(* IEC 61131-3 sources: model-first-plc-agent-ai/results/T3-B-12, 1 file *)

(* ---- b_code.st ---- *)
FUNCTION_BLOCK FillingTankControl
VAR_INPUT
    start : BOOL;
    stop : BOOL;
    LSH : BOOL;
    LSHH : BOOL;
    TON_Duration : TIME;
    TOF_Duration : TIME;
END_VAR
VAR_OUTPUT
    fill_valve : BOOL;
    discharge_valve : BOOL;
END_VAR
VAR
    state_id : INT := 0;
    filling_active : BOOL;
    ton_q : BOOL;
    tof_q : BOOL;
    fill_timer : TON;
    pause_timer : TOF;
END_VAR

(* States: 0 = idle, 1 = filling, 2 = pause. *)
(* Both level switches inhibit filling; LSHH is a safety override. *)
IF stop OR LSH OR LSHH THEN
    state_id := 0;
ELSIF (state_id = 0) AND start THEN
    state_id := 1;
END_IF;

filling_active := (state_id = 1);

fill_timer(
    IN := filling_active,
    PT := TON_Duration
);
ton_q := fill_timer.Q;

pause_timer(
    IN := filling_active,
    PT := TOF_Duration
);
tof_q := pause_timer.Q;

IF NOT (stop OR LSH OR LSHH) THEN
    CASE state_id OF
        0:
            state_id := 0;

        1:
            IF ton_q THEN
                state_id := 2;
            END_IF;

        2:
            IF NOT tof_q THEN
                state_id := 1;
            END_IF;

        ELSE
            state_id := 0;
    END_CASE;
END_IF;

fill_valve := (state_id = 1) AND NOT stop AND NOT LSH AND NOT LSHH;
discharge_valve := FALSE;

END_FUNCTION_BLOCK

PROGRAM Main
VAR
    StartCommand AT %IX100.0 : BOOL;
    StopCommand AT %IX100.1 : BOOL;
    LSH AT %IX100.2 : BOOL;
    LSHH AT %IX100.3 : BOOL;
    FillValve AT %QX100.0 : BOOL;
    DischargeValve AT %QX100.1 : BOOL;
END_VAR
VAR
    (* Adjustable timer parameters; these are initial defaults. *)
    TON_Duration : TIME := T#5s;
    TOF_Duration : TIME := T#2s;

    start : BOOL;
    stop : BOOL;
    start_edge : R_TRIG;
    tank_control : FillingTankControl;
END_VAR

start_edge(CLK := StartCommand);
start := start_edge.Q;
stop := StopCommand;

tank_control(
    start := start,
    stop := stop,
    LSH := LSH,
    LSHH := LSHH,
    TON_Duration := TON_Duration,
    TOF_Duration := TOF_Duration
);

FillValve := tank_control.fill_valve;
DischargeValve := tank_control.discharge_valve;

END_PROGRAM
